(* IEC 61131-3 sources: SemantiST/compiler/intake/normalize/probes/scl-begin, 2 files *)

(* ---- original.st ---- *)
FUNCTION INC : INT
VAR_INPUT
    X : INT;
END_VAR
BEGIN
INC := X + 1;
END_FUNCTION

FUNCTION main : DINT
printf('%d$N', INC(10));
main := 0;
END_FUNCTION

(* ---- rewritten.st ---- *)
FUNCTION INC : INT
VAR_INPUT
    X : INT;
END_VAR
(* BEGIN *)
INC := X + 1;
END_FUNCTION

FUNCTION main : DINT
printf('%d$N', INC(10));
main := 0;
END_FUNCTION
